{region 'Documentation'}
(*!
<summary>Run Control request and status view; the execution owner calls the concrete FB cyclically.</summary>
<description>
Request methods record same-task intent; they do not execute the lifecycle synchronously. Repeated requests coalesce and regular processing applies Reset over Abort over Start. Status is a stored value snapshot. Name and Result are inherited from I_ResultProvider. The concrete owner must still be called cyclically, including after completion.
</description>
*)
{endregion}
INTERFACE I_RunControl EXTENDS I_ResultProvider

{region 'Documentation'}
(*!
<summary>Records an abort request for regular lifecycle processing.</summary>
*)
{endregion}
METHOD RequestAbort
END_METHOD

{region 'Documentation'}
(*!
<summary>Records a reset request for regular lifecycle processing.</summary>
*)
{endregion}
METHOD RequestReset
END_METHOD

{region 'Documentation'}
(*!
<summary>Records a start request for regular lifecycle processing.</summary>
*)
{endregion}
METHOD RequestStart
END_METHOD

{region 'Documentation'}
(*!
<summary>Current owner status snapshot; reading does not execute lifecycle processing.</summary>
*)
{endregion}
PROPERTY Status : ST_RunControlStatus //! Current owner status snapshot; reading does not execute lifecycle processing.
GET // PUBLIC
END_GET
END_PROPERTY

END_INTERFACE

(* stored: Version 1.1.0.1
   Itf I_RunControl: Id {da624c3d-f407-4da3-bfdc-c101fd2b858f}
   Method RequestAbort: Id {31ac04f8-4a29-444c-9ae6-375550190ddc}
   Method RequestReset: Id {933c2d85-a2c5-4aa2-b523-f50804b414f7}
   Method RequestStart: Id {0e4bdb41-5fee-4d72-a83c-4fe8092b7b76}
   Property Status: Id {380f3aef-f890-43e9-b0cc-1aad8b1538bc}
   Get Get: Id {beff11d8-6078-4cc7-b4e4-22a804dde9f1} *)
